(* IEC 61131-3 sources: Automatic-Tank-Level-and-Pump-Control-System/tankmanualAuto/pous/programs, 1 file *)

(* ---- main.st ---- *)
PROGRAM main
  VAR
    START : BOOL;
    STOP : BOOL;
    AUTO_MODE : BOOL;
    PUMP_RUN_FEEDBACK : BOOL;
    OVERLOAD_TRIP : BOOL;
    STARTUP_TIMER : TON;
    START_FAILURE : BOOL;
    MANUAL_MODE : BOOL;
    TANK_LEVEL : REAL;
    PUMP : BOOL;
    MANUAL_START : BOOL;
    MANUAL_STOP : BOOL;
    SYSTEM_RUN : BOOL;
    auto_select : BOOL;
    manual_select : BOOL;
    level_real : DINT;
    sensor_fault : BOOL;
    alarm_light_red : BOOL;
    sensor_fault_latched : BOOL;
    sensor_reset : BOOL;
    START_FAILURE_RESET : BOOL;
    PUMP_FAULT_ALARM : BOOL;
    OVERLOAD_FAULT_LATCHED : BOOL;
    OVERLOAD_RESET : BOOL;
  END_VAR

if STOP then
    SYSTEM_RUN:= false;
elsif START then
     SYSTEM_RUN:= true;
end_if;

IF (level_real < 0) OR (level_real > 32767) THEN
    SENSOR_FAULT_LATCHED := TRUE;
END_IF;

IF sensor_reset AND (level_real >= 0) AND (level_real <= 32767) THEN
    SENSOR_FAULT_LATCHED := FALSE;
END_IF;

sensor_fault := SENSOR_FAULT_LATCHED;

IF sensor_fault THEN
    TANK_LEVEL := -1.0;
    alarm_light_red := TRUE;
ELSE
    TANK_LEVEL := DINT_TO_REAL(level_real) * 100.0 / 32767.0;
    alarm_light_red := FALSE;
END_IF;

IF AUTO_SELECT AND NOT MANUAL_SELECT THEN
    AUTO_MODE := TRUE;
    MANUAL_MODE := FALSE;

ELSIF MANUAL_SELECT AND NOT AUTO_SELECT THEN
    MANUAL_MODE := TRUE;
    AUTO_MODE := FALSE;

ELSIF AUTO_SELECT AND MANUAL_SELECT THEN
    AUTO_MODE := FALSE;
    MANUAL_MODE := FALSE;
END_IF;

IF NOT SYSTEM_RUN THEN
    PUMP := FALSE;
ELSIF sensor_fault THEN
    PUMP := FALSE;

ELSIF AUTO_MODE THEN
    IF TANK_LEVEL <= 30.0 THEN
        PUMP := TRUE;
    ELSIF TANK_LEVEL >= 90.0 THEN
        PUMP := FALSE;
    END_IF;

ELSIF MANUAL_MODE THEN
    IF MANUAL_STOP THEN
        PUMP := FALSE;
    ELSIF MANUAL_START THEN
        PUMP := TRUE;
    END_IF;

ELSE
    PUMP := FALSE;
END_IF;

STARTUP_TIMER (
    IN := PUMP AND NOT PUMP_RUN_FEEDBACK,
    PT := T#3s
);
IF STARTUP_TIMER.Q THEN
    START_FAILURE := TRUE;
END_IF;

IF START_FAILURE_RESET
   AND NOT PUMP
   AND NOT PUMP_RUN_FEEDBACK
   AND NOT OVERLOAD_TRIP
   AND NOT sensor_fault THEN

    START_FAILURE := FALSE;
END_IF;

PUMP_FAULT_ALARM := START_FAILURE OR OVERLOAD_FAULT_LATCHED;

IF sensor_fault OR OVERLOAD_FAULT_LATCHED OR START_FAILURE THEN
    PUMP := FALSE;
END_IF;
IF OVERLOAD_TRIP THEN
    OVERLOAD_FAULT_LATCHED := TRUE;
END_IF;

IF OVERLOAD_TRIP THEN
    OVERLOAD_FAULT_LATCHED := TRUE;
END_IF;

IF OVERLOAD_RESET
   AND NOT OVERLOAD_TRIP
   AND NOT PUMP
   AND NOT PUMP_RUN_FEEDBACK THEN

    OVERLOAD_FAULT_LATCHED := FALSE;
END_IF;

END_PROGRAM
